TYPE HardwareError :
STRUCT
	isActive : BOOL;
	id : UDINT;
	text : STRING(80);
END_STRUCT
END_TYPE

(* stored: Version 1.1.0.1, ProductVersion 3.1.4026.12
   DUT HardwareError: Id {5b37c64c-1c38-5faf-a768-5ff4e757a912} *)
